{attribute 'TcGenerated'}
{attribute 'no-analysis'}
{attribute 'linkalways'}
// This function has been automatically generated from the project information.
VAR_GLOBAL CONSTANT
	{attribute 'const_non_replaced'}
	stLibVersion_LPLC : ST_LibVersion := (iMajor := 2, iMinor := 2, iBuild := 0, iRevision := 0, nFlags := 0, sVersion := '2.2.0');
END_VAR

(* stored: Version 1.1.0.1
   GVL Global_Version: Id {3579d7a9-aa55-4461-9b4a-a7719b763321} *)
